// TwinCAT 3 PLC project PLCSim
// ProgramVersion: 3.1.4026.20
// libraries:
//   Tc2_Standard, * (Beckhoff Automation GmbH)
//   Tc2_System, * (Beckhoff Automation GmbH)
//   Tc3_Module, * (Beckhoff Automation GmbH)
//   VisuDialogs, * (System)
// project tree:
//   / GlobalTextList.TcGTLO, PlcTask.TcTTO, Visualization Manager.TcVMO (not stored)
//   GVLs/ GVL.TcGVL
//   POUs/ MAIN.TcPOU
//   VISUs/ Visualization.TcVIS
// real-time tasks:
//   TASK PlcTask: cycle T#10ms, priority 20, ADS port 350
// variable links:
//   PLCSim/PLCSim Instance <-> PLCStudent/PLCStudent Instance
//     PlcTask Inputs/GVL.ixLed{1..8} <-> PlcTask Outputs/ControlFBD.qxLed{1..8}  (8 links)
//     PlcTask Outputs/GVL.qxButton{1..8} <-> PlcTask Inputs/ControlFBD.ixButton{1..8}  (8 links)

CONFIGURATION PLCSim
    RESOURCE PLC ON TwinCAT3
        TASK PlcTask(INTERVAL := T#10ms, PRIORITY := 20);
        PROGRAM MAIN WITH PlcTask : MAIN;
    END_RESOURCE
END_CONFIGURATION

// ---- GVLs/GVL.TcGVL
{attribute 'qualified_only'}
VAR_GLOBAL
	qxButton1 AT %Q* : BOOL;
	qxButton2 AT %Q* : BOOL;
	qxButton3 AT %Q* : BOOL;
	qxButton4 AT %Q* : BOOL;
	qxButton5 AT %Q* : BOOL;
	qxButton6 AT %Q* : BOOL;
	qxButton7 AT %Q* : BOOL;
	qxButton8 AT %Q* : BOOL;
	
	ixLed1 AT %I* : BOOL;
	ixLed2 AT %I* : BOOL;
	ixLed3 AT %I* : BOOL;
	ixLed4 AT %I* : BOOL;
	ixLed5 AT %I* : BOOL;
	ixLed6 AT %I* : BOOL;
	ixLed7 AT %I* : BOOL;
	ixLed8 AT %I* : BOOL;
END_VAR

// ---- POUs/MAIN.TcPOU
PROGRAM MAIN
VAR
END_VAR

END_PROGRAM

// ---- GlobalTextList.TcGTLO
TEXTLIST GlobalTextList
  308 = '1              2             3             4             5              6             7             8'
  309 = 'Connector IN'
  310 = 'Connector OUT'
  306 = 'I/O Box'
  307 = 'University West \nAnders N Dec 2018'
END_TEXTLIST

// ---- VISUs/Visualization.TcVIS
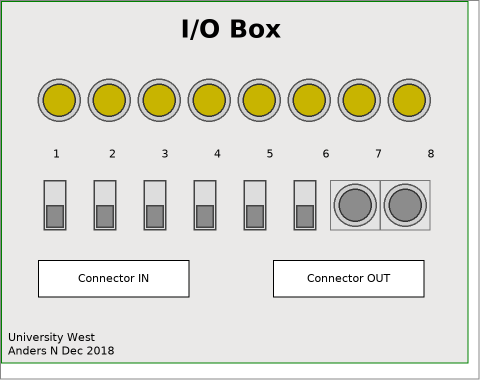
VISUALIZATION Visualization  // 480x380
    Rectangle (1,1 467x362)
    Label (147,0 168x57), "I/O Box"
    Lamp1 (34,75 50x50), variable: GVL.ixLed1, style: Lamp-Lamp1-Yellow
    Lamp1 (84,75 50x50), variable: GVL.ixLed2, style: Lamp-Lamp1-Yellow
    Lamp1 (134,75 50x50), variable: GVL.ixLed3, style: Lamp-Lamp1-Yellow
    Lamp1 (184,75 50x50), variable: GVL.ixLed4, style: Lamp-Lamp1-Yellow
    Lamp1 (234,75 50x50), variable: GVL.ixLed5, style: Lamp-Lamp1-Yellow
    Lamp1 (284,75 50x50), variable: GVL.ixLed6, style: Lamp-Lamp1-Yellow
    Lamp1 (334,75 50x50), variable: GVL.ixLed7, style: Lamp-Lamp1-Yellow
    Lamp1 (384,75 50x50), variable: GVL.ixLed8, style: Lamp-Lamp1-Yellow
    Label (5,329 118x30), "University West Anders N Dec 2018"
    Label (50,144 392x20), "1 2 3 4 5 6 7 8"
    RoundedRectangle (38,260 151x37), "Connector IN"
    RoundedRectangle (273,260 151x37), "Connector OUT"
    DipSwitch (30,180 50x50), variable: GVL.qxButton1, behaviour: TOGGLE, style: Switch-DipSwitch-Gray
    DipSwitch (80,180 50x50), variable: GVL.qxButton2, behaviour: TOGGLE, style: Switch-DipSwitch-Gray
    DipSwitch (130,180 50x50), variable: GVL.qxButton3, behaviour: TOGGLE, style: Switch-DipSwitch-Gray
    DipSwitch (180,180 50x50), variable: GVL.qxButton4, behaviour: TOGGLE, style: Switch-DipSwitch-Gray
    DipSwitch (230,180 50x50), variable: GVL.qxButton5, behaviour: TOGGLE, style: Switch-DipSwitch-Gray
    DipSwitch (280,180 50x50), variable: GVL.qxButton6, behaviour: TOGGLE, style: Switch-DipSwitch-Gray
    PushSwitch (330,180 50x50), variable: GVL.qxButton7, behaviour: TAP, style: Switch-PushSwitch-Gray
    PushSwitch (380,180 50x50), variable: GVL.qxButton8, behaviour: TAP, style: Switch-PushSwitch-Gray
    hotkey HotkeyInput Id=481044725760, Key=KeyName=1, VisuElemId=-1
END_VISUALIZATION
